// TIA Portal V20 export
Screen "Pop-up_USER_OPERATION_LEGEND_Popup"  380x350
  ScreenItem "Background" at 0,0 size 380x350  Type=HmiRectangle
  ScreenItem "Textfeld_9" at 223,315 size 126x20  Type=HmiTextBox
  ScreenItem "Textfeld_Legende" at 1,1 size 378x45  Type=HmiTextBox
  ScreenItem "Textfeld_15" at 10,50 size 305x30  Type=HmiTextBox
  ScreenItem "Textfeld_17" at 10,88 size 66x20  Type=HmiTextBox
  ScreenItem "PB_ADV" at 137,111 size 46x31  Type=HmiButton
  ScreenItem "PB_RTN" at 235,110 size 46x31  Type=HmiButton
  ScreenItem "ADV_Slow" at 128,178 size 62x18  Type=HmiButton
  ScreenItem "Textfeld_1" at 142,82 size 60x30  Type=HmiTextBox
  ScreenItem "Textfeld_2" at 238,82 size 60x30  Type=HmiTextBox
  ScreenItem "Textfeld_3" at 10,147 size 66x20  Type=HmiTextBox
  ScreenItem "ADV_Slow_1" at 229,178 size 62x18  Type=HmiButton
  ScreenItem "Textfeld_4" at 10,177 size 66x20  Type=HmiTextBox
  ScreenItem "ADV_Slow_2" at 128,206 size 62x18  Type=HmiButton
  ScreenItem "ADV_Slow_3" at 229,206 size 62x18  Type=HmiButton
  ScreenItem "Textfeld_5" at 10,206 size 104x20  Type=HmiTextBox
  ScreenItem "Textfeld_6" at 10,254 size 66x20  Type=HmiTextBox
  ScreenItem "ADV_Slow_4" at 125,254 size 62x18  Type=HmiButton
  ScreenItem "ADV_Slow_5" at 124,284 size 62x18  Type=HmiButton
  ScreenItem "Textfeld_7" at 226,253 size 105x20  Type=HmiTextBox
  ScreenItem "Textfeld_8" at 223,282 size 126x20  Type=HmiTextBox
  ScreenItem "PB_ADV_1" at 133,314 size 46x31  Type=HmiButton
  ScreenItem "Cancel Mode" at 289,1 size 90x60  Type=HmiButton
